FUNCTION VC_GetInt8 : SINT
// Reads Int8 (1 byte, little-endian) from Buf[Pos] and advances Pos.
VAR_IN_OUT
    Buf   : ARRAY[*] OF BYTE;
    Pos   : UDINT;
END_VAR
VAR
    nVal : SINT;
END_VAR

nVal := 0;
VC_GetRaw(Buf := Buf, Pos := Pos, pDst := ADR(nVal), Size := 1);
VC_GetInt8 := nVal;

END_FUNCTION

(* stored: Version 1.1.0.1, ProductVersion 3.1.4024.12
   POU VC_GetInt8: Id {f5fdc942-f272-426e-8fc3-2911677a06d4}, SpecialFunc None *)
